RoboDK station: PickPlace_Delta_Fanuc.rdk

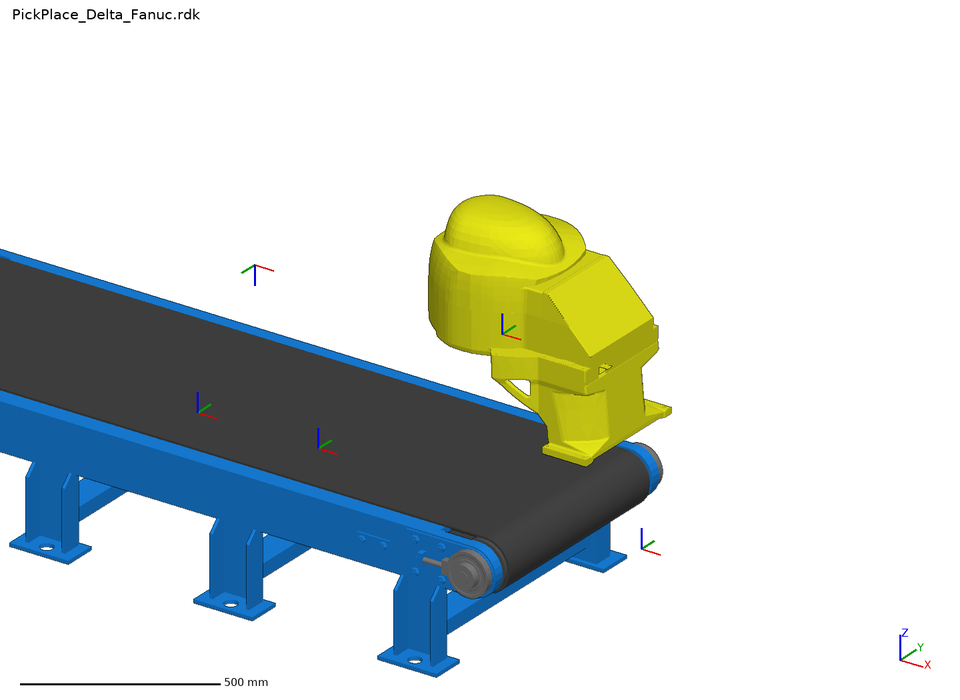
[picture v0: the station drawn from its stored meshes, robots at their saved joint values, targets as dots, program paths as lines]
Station PickPlace_Delta_Fanuc (saved by RoboDK 6.0.1). Poses are relative to the parent item; angles as X-Y-Z fixed-axis rotations.
Station parameters (name, value as stored): SICK WL4S Laser Sensor, 0, start_prox, 0
  - frame Conveyor Belt Wide (2m) Base at (0, 0, 0) mm
    - robot Conveyor Belt Wide (2m): 1 axes
        modified DH rows (alpha deg, a mm, theta deg, d mm): 0, 0, 0, 0 linear
        base shift (0, 0, 0) mm, rotated rx 0 ry 90 rz 0 deg
        joint limits [-900000] to [900000]; home [0]; saved at [-467637]
      - frame Conveyor Frame at (0, 0, 0) mm
        - object Box at (476786, 176.94, 12.44) mm, rotated rx -0.58 ry 0.13 rz -5.1 deg, size 10 x 20 x 5 mm, geometry from box.sld
        - object Box at (476618, 129.49, 12.91) mm, rotated rx -0.57 ry 0.15 rz -3.3 deg, size 10 x 20 x 5 mm, geometry from box.sld
        - object Box at (476349, 147.41, 12.73) mm, rotated rx -0.57 ry 0.15 rz -3.78 deg, size 10 x 20 x 5 mm, geometry from box.sld
        - object Box at (476190, 165.56, 12.56) mm, rotated rx -0.58 ry 0.12 rz -6.59 deg, size 10 x 20 x 5 mm, geometry from box.sld
        - object Box at (476046, 14.84, 14.04) mm, rotated rx -0.54 ry 0.25 rz 6.85 deg, size 10 x 20 x 5 mm, geometry from box.sld
        - object Box at (475925, 101.99, 13.18) mm, rotated rx -0.51 ry 0.3 rz 12.4 deg, size 10 x 20 x 5 mm, geometry from box.sld
        - object Box at (475776, 10.76, 14.08) mm, rotated rx -0.59 ry 0.06 rz -12.55 deg, size 10 x 20 x 5 mm, geometry from box.sld
        - object Box at (475609, 201.57, 12.2) mm, rotated rx -0.51 ry 0.3 rz 12.73 deg, size 10 x 20 x 5 mm, geometry from box.sld
        - object Box at (475416, 151.6, 12.69) mm, rotated rx -0.58 ry 0.11 rz -7.36 deg, size 10 x 20 x 5 mm, geometry from box.sld
        - object Box at (475210, 21.91, 13.97) mm, rotated rx -0.59 ry 0.1 rz -8.46 deg, size 10 x 20 x 5 mm, geometry from box.sld
        - object Box at (475016, 87.28, 13.33) mm, rotated rx -0.59 ry 0.08 rz -10.47 deg, size 10 x 20 x 5 mm, geometry from box.sld
        - object Box at (474824, 137.82, 12.83) mm, rotated rx -0.51 ry 0.31 rz 12.89 deg, size 10 x 20 x 5 mm, geometry from box.sld
        - object Box at (474629, 180.76, 12.41) mm, rotated rx -0.55 ry 0.21 rz 2.74 deg, size 10 x 20 x 5 mm, geometry from box.sld
        - object Box at (474453, 158.14, 12.63) mm, rotated rx -0.53 ry 0.27 rz 8.81 deg, size 10 x 20 x 5 mm, geometry from box.sld
        - object Box at (474289, 158.23, 12.63) mm, rotated rx -0.54 ry 0.25 rz 7.11 deg, size 10 x 20 x 5 mm, geometry from box.sld
    - frame Reference Box Frame at (60, 290, 366.5) mm
      - object ref_obj at (0, 0, 0) mm, size 252 x 305.4 x 216.7 mm, geometry from Box-12x10in-Closed.sld
      - object ref_lid at (-60, -186.65, 13.17) mm, rotated rx -0.56 ry 0.19 rz 0 deg, size 10 x 20 x 5 mm, geometry from box.sld
    - object SICK WL4S Laser Sensor at (1954, -20, 370) mm, rotated rx 180 ry 0 rz 90 deg, size 683.3 x 45.2 x 12.5 mm, geometry from SICK-WL4S-Laser-Sensor.sld
    - object start_prox at (0, -20, 370) mm, rotated rx 180 ry 0 rz 90 deg, size 683.3 x 45.2 x 12.5 mm, geometry from SICK-WL4S-Laser-Sensor.sld
  - program MainProgram (5 instructions, listed below)
  - notes Description: <!DOCTYPE HTML PUBLIC "-//W3C//DTD HTML 4.0//EN" "http://www.w3.org/TR/REC-html40/strict.dtd">
<html><head><meta name="qrichtext" content="1" /><style type="text/css">
p, li { white-space: pre-wrap; }
</style></head><body style=" font-family:'MS Shell Dlg 2'; font-size:8.25pt; font-weight:400; font-style:normal;">
<p style=" margin-top:0px; margin-bottom:0px; margin-left:0px; margin-right:0px; -qt-block-indent:0; text-indent:0px;">This example demonstrates a conveyor simulation in RoboDK using Python scripting. A script generates boxes of varying sizes and positions while the conveyor moves continuously. A sensor detects when a box reaches the conveyor’s edge and stops the conveyor. The station showcases how conveyors, part generation, and sensor-based control can be simulated with the API.</p></body></html>
  - frame Fanuc M-1iA/0.5SL Base at (1954.3, 143.51, 858.22) mm
    - robot Fanuc M-1iA/0.5SL: 4 axes, payload 0.5 kg, reach 420 mm, repeatability 0.03 mm, weight 23 kg
        joint limits [-25, -25, -25, -36000] to [80, 80, 80, 36000]; home [0, 0, 0, 0]; saved at [8.958, 51.399, -22.511, 0]
      - tool Tool 1, TCP at (0, 0, 0) mm
        - object Box at (56.03, -11.25, -8.71) mm, rotated rx 179.51 ry -0.34 rz -16.22 deg, size 10 x 20 x 5 mm, geometry from box.sld
  - frame CamFrame at (1207.08, 136.9, 843.5) mm, rotated rx -180 ry -0.2 rz -0.44 deg
    - camera Camera 1
  - frame Frame 6 at (1375.31, 171.47, 367.78) mm
  - frame Frame 7 at (1050, 111.47, 400) mm
  - frame delete_box_frame at (2400, 111.47, 400) mm

--- program MainProgram (robot Conveyor Belt Wide (2m)) ---
  Call ConveyorReset
  Run SensorReader
  Set speed (25.0 mm/s)
  Run ConveyorRunner
  Run BoxSpawner
